Staubli VAL3: init.pgx

program init()
begin
  _nClock=0
  call io:init()
end
